(* IEC 61131-3 sources: plc-st-coding-agent/progress/f14_candidate/release/review/fixtures/agent_9772562, 4 files *)

(* ---- arm_one_step.st ---- *)
FUNCTION_BLOCK FB
VAR_INPUT
    ManualMode : BOOL;
    SingleStepMode : BOOL;
    SingleCycleMode : BOOL;
    ContinuousMode : BOOL;
    EmergencyStop : BOOL;
    Start : BOOL;
    DownButton : BOOL;
    UpButton : BOOL;
    LeftButton : BOOL;
    RightButton : BOOL;
    GripButton : BOOL;
    ReleaseButton : BOOL;
    DownLimitSwitch : BOOL;
    UpLimitSwitch : BOOL;
    LeftLimitSwitch : BOOL;
    RightLimitSwitch : BOOL;
    GripLimitSwitch : BOOL;
    ReleaseLimitSwitch : BOOL;
END_VAR
VAR_OUTPUT
    MoveDown : BOOL;
    MoveUp : BOOL;
    MoveLeft : BOOL;
    MoveRight : BOOL;
    ActivateGrip : BOOL;
    ActivateRelease : BOOL;
END_VAR
VAR
    step : INT := 1;
    busy : BOOL := FALSE;
    prevStart : BOOL := FALSE;
    prevManual : BOOL := FALSE;
    prevSingleStep : BOOL := FALSE;
    prevSingleCycle : BOOL := FALSE;
    prevContinuous : BOOL := FALSE;
    startRising : BOOL;
    autoSelected : BOOL;
    stepDone : BOOL;
END_VAR

(* 模式变化检测：任何模式输入改变时，停止当前动作并复位步骤 *)
IF (ManualMode <> prevManual) OR (SingleStepMode <> prevSingleStep) OR (SingleCycleMode <> prevSingleCycle) OR (ContinuousMode <> prevContinuous) THEN
    busy := FALSE;
    step := 1;
END_IF;
prevManual := ManualMode;
prevSingleStep := SingleStepMode;
prevSingleCycle := SingleCycleMode;
prevContinuous := ContinuousMode;

autoSelected := NOT ManualMode AND (SingleStepMode OR SingleCycleMode OR ContinuousMode);

startRising := Start AND NOT prevStart;
prevStart := Start;

IF autoSelected AND EmergencyStop THEN
    IF startRising THEN
        IF NOT busy THEN
            busy := TRUE;
        END_IF;
    END_IF;

    IF busy THEN
        stepDone := FALSE;
        CASE step OF
            1: stepDone := DownLimitSwitch;
            2: stepDone := GripLimitSwitch;
            3: stepDone := UpLimitSwitch;
            4: stepDone := RightLimitSwitch;
            5: stepDone := DownLimitSwitch;
            6: stepDone := ReleaseLimitSwitch;
            7: stepDone := UpLimitSwitch;
            8: stepDone := LeftLimitSwitch;
        END_CASE;

        IF stepDone THEN
            IF SingleStepMode THEN
                busy := FALSE;
                step := step MOD 8 + 1;
            ELSIF SingleCycleMode THEN
                IF step = 8 THEN
                    busy := FALSE;
                    step := 1;
                ELSE
                    step := step + 1;
                END_IF;
            ELSIF ContinuousMode THEN
                step := step MOD 8 + 1;
            END_IF;
        END_IF;
    END_IF;
END_IF;

IF EmergencyStop THEN
    IF ManualMode THEN
        MoveDown := DownButton AND NOT UpButton AND NOT DownLimitSwitch;
        MoveUp := UpButton AND NOT DownButton AND NOT UpLimitSwitch;
        MoveLeft := LeftButton AND NOT RightButton AND NOT LeftLimitSwitch;
        MoveRight := RightButton AND NOT LeftButton AND NOT RightLimitSwitch;
        ActivateGrip := GripButton AND NOT ReleaseButton AND NOT GripLimitSwitch;
        ActivateRelease := ReleaseButton AND NOT GripButton AND NOT ReleaseLimitSwitch;
    ELSIF autoSelected THEN
        IF busy THEN
            MoveDown := ((step = 1) OR (step = 5)) AND NOT DownLimitSwitch;
            MoveUp := ((step = 3) OR (step = 7)) AND NOT UpLimitSwitch;
            MoveLeft := (step = 8) AND NOT LeftLimitSwitch;
            MoveRight := (step = 4) AND NOT RightLimitSwitch;
            ActivateGrip := (step = 2) AND NOT GripLimitSwitch;
            ActivateRelease := (step = 6) AND NOT ReleaseLimitSwitch;
        ELSE
            MoveDown := FALSE;
            MoveUp := FALSE;
            MoveLeft := FALSE;
            MoveRight := FALSE;
            ActivateGrip := FALSE;
            ActivateRelease := FALSE;
        END_IF;
    ELSE
        MoveDown := FALSE;
        MoveUp := FALSE;
        MoveLeft := FALSE;
        MoveRight := FALSE;
        ActivateGrip := FALSE;
        ActivateRelease := FALSE;
    END_IF;
ELSE
    MoveDown := FALSE;
    MoveUp := FALSE;
    MoveLeft := FALSE;
    MoveRight := FALSE;
    ActivateGrip := FALSE;
    ActivateRelease := FALSE;
END_IF;

END_FUNCTION_BLOCK

(* ---- arm_restart.st ---- *)
FUNCTION_BLOCK FB
VAR_INPUT
    ManualMode : BOOL;
    SingleStepMode : BOOL;
    SingleCycleMode : BOOL;
    ContinuousMode : BOOL;
    EmergencyStop : BOOL;
    Start : BOOL;
    DownButton : BOOL;
    UpButton : BOOL;
    LeftButton : BOOL;
    RightButton : BOOL;
    GripButton : BOOL;
    ReleaseButton : BOOL;
    DownLimitSwitch : BOOL;
    UpLimitSwitch : BOOL;
    LeftLimitSwitch : BOOL;
    RightLimitSwitch : BOOL;
    GripLimitSwitch : BOOL;
    ReleaseLimitSwitch : BOOL;
END_VAR
VAR_OUTPUT
    MoveDown : BOOL;
    MoveUp : BOOL;
    MoveLeft : BOOL;
    MoveRight : BOOL;
    ActivateGrip : BOOL;
    ActivateRelease : BOOL;
END_VAR
VAR
    StartPrev : BOOL := FALSE;
    PrevManualMode : BOOL := FALSE;
    PrevSingleStepMode : BOOL := FALSE;
    PrevSingleCycleMode : BOOL := FALSE;
    PrevContinuousMode : BOOL := FALSE;
    ModeChanged : BOOL;
    StartPulse : BOOL;
    AutoStep : INT := 0;
END_VAR

MoveDown := FALSE;
MoveUp := FALSE;
MoveLeft := FALSE;
MoveRight := FALSE;
ActivateGrip := FALSE;
ActivateRelease := FALSE;

StartPulse := Start AND NOT StartPrev;
ModeChanged := (ManualMode <> PrevManualMode)
                OR (SingleStepMode <> PrevSingleStepMode)
                OR (SingleCycleMode <> PrevSingleCycleMode)
                OR (ContinuousMode <> PrevContinuousMode);

IF ModeChanged THEN
    AutoStep := 0;
END_IF;

IF EmergencyStop THEN
    IF ManualMode THEN
        MoveDown := DownButton AND NOT UpButton AND NOT DownLimitSwitch;
        MoveUp := UpButton AND NOT DownButton AND NOT UpLimitSwitch;
        MoveLeft := LeftButton AND NOT RightButton AND NOT LeftLimitSwitch;
        MoveRight := RightButton AND NOT LeftButton AND NOT RightLimitSwitch;
        ActivateGrip := GripButton AND NOT ReleaseButton AND NOT GripLimitSwitch;
        ActivateRelease := ReleaseButton AND NOT GripButton AND NOT ReleaseLimitSwitch;
    ELSIF SingleStepMode THEN
        IF AutoStep = 0 THEN
            IF StartPulse THEN
                AutoStep := 1;
            END_IF;
        END_IF;

        CASE AutoStep OF
            1:
                IF DownLimitSwitch THEN
                    AutoStep := 0;
                ELSE
                    MoveDown := TRUE;
                END_IF;
            2:
                IF GripLimitSwitch THEN
                    AutoStep := 0;
                ELSE
                    ActivateGrip := TRUE;
                END_IF;
            3:
                IF UpLimitSwitch THEN
                    AutoStep := 0;
                ELSE
                    MoveUp := TRUE;
                END_IF;
            4:
                IF RightLimitSwitch THEN
                    AutoStep := 0;
                ELSE
                    MoveRight := TRUE;
                END_IF;
            5:
                IF DownLimitSwitch THEN
                    AutoStep := 0;
                ELSE
                    MoveDown := TRUE;
                END_IF;
            6:
                IF ReleaseLimitSwitch THEN
                    AutoStep := 0;
                ELSE
                    ActivateRelease := TRUE;
                END_IF;
            7:
                IF UpLimitSwitch THEN
                    AutoStep := 0;
                ELSE
                    MoveUp := TRUE;
                END_IF;
            8:
                IF LeftLimitSwitch THEN
                    AutoStep := 0;
                ELSE
                    MoveLeft := TRUE;
                END_IF;
        END_CASE;
    ELSIF SingleCycleMode OR ContinuousMode THEN
        IF AutoStep = 0 THEN
            IF StartPulse THEN
                AutoStep := 1;
            END_IF;
        END_IF;

        IF AutoStep = 1 AND DownLimitSwitch THEN
            AutoStep := 2;
        END_IF;
        IF AutoStep = 2 AND GripLimitSwitch THEN
            AutoStep := 3;
        END_IF;
        IF AutoStep = 3 AND UpLimitSwitch THEN
            AutoStep := 4;
        END_IF;
        IF AutoStep = 4 AND RightLimitSwitch THEN
            AutoStep := 5;
        END_IF;
        IF AutoStep = 5 AND DownLimitSwitch THEN
            AutoStep := 6;
        END_IF;
        IF AutoStep = 6 AND ReleaseLimitSwitch THEN
            AutoStep := 7;
        END_IF;
        IF AutoStep = 7 AND UpLimitSwitch THEN
            AutoStep := 8;
        END_IF;
        IF AutoStep = 8 AND LeftLimitSwitch THEN
            IF ContinuousMode THEN
                AutoStep := 1;
            ELSE
                AutoStep := 0;
            END_IF;
        END_IF;

        CASE AutoStep OF
            1:
                IF NOT DownLimitSwitch THEN
                    MoveDown := TRUE;
                END_IF;
            2:
                IF NOT GripLimitSwitch THEN
                    ActivateGrip := TRUE;
                END_IF;
            3:
                IF NOT UpLimitSwitch THEN
                    MoveUp := TRUE;
                END_IF;
            4:
                IF NOT RightLimitSwitch THEN
                    MoveRight := TRUE;
                END_IF;
            5:
                IF NOT DownLimitSwitch THEN
                    MoveDown := TRUE;
                END_IF;
            6:
                IF NOT ReleaseLimitSwitch THEN
                    ActivateRelease := TRUE;
                END_IF;
            7:
                IF NOT UpLimitSwitch THEN
                    MoveUp := TRUE;
                END_IF;
            8:
                IF NOT LeftLimitSwitch THEN
                    MoveLeft := TRUE;
                END_IF;
        END_CASE;
    END_IF;
END_IF;

PrevManualMode := ManualMode;
PrevSingleStepMode := SingleStepMode;
PrevSingleCycleMode := SingleCycleMode;
PrevContinuousMode := ContinuousMode;
StartPrev := Start;
END_FUNCTION_BLOCK

(* ---- conveyor.st ---- *)
FUNCTION_BLOCK FB
VAR_INPUT
    processLength : USINT;
    sensor1 : BOOL;
    sensor2 : BOOL;
    sensor3 : BOOL;
    sensor4 : BOOL;
    sensor5 : BOOL;
    station1Start : BOOL;
    station2Complete : BOOL;
    station3Complete : BOOL;
    station4Complete : BOOL;
    processSequence : ARRAY[1..8] OF USINT;
END_VAR
VAR_OUTPUT
    conveyorLeft : BOOL;
    conveyorRight : BOOL;
END_VAR
VAR
    state : USINT := 0; (* 0=IDLE, 1=MOVING, 2=WAIT_PROCESS, 3=DONE *)
    currentStation : USINT := 1;
    seqIndex : USINT := 1;
    targetStation : USINT := 5;
    lastStation1Start : BOOL := FALSE;
    lastComplete2 : BOOL := FALSE;
    lastComplete3 : BOOL := FALSE;
    lastComplete4 : BOOL := FALSE;
END_VAR

(* 默认输出 *)
conveyorLeft := FALSE;
conveyorRight := FALSE;

(* 检查 processLength 有效性：若无效则强制停止并保持初始状态 *)
IF (processLength < 1) OR (processLength > 8) THEN
    state := 0;
    currentStation := 1;
    seqIndex := 1;
ELSE
    (* 状态机 *)
    IF (state = 0) OR (state = 3) THEN
        (* 启动检测：1# 传感器有料且启动按钮上升沿 *)
        IF (NOT lastStation1Start) AND station1Start AND sensor1 THEN
            seqIndex := 1;
            currentStation := 1;
            targetStation := processSequence[1];
            state := 1; (* MOVING *)
        END_IF
    ELSIF state = 1 THEN
        (* 移动中，检测目标传感器 *)
        IF (targetStation = 2) AND sensor2 THEN
            currentStation := 2;
            IF targetStation = 5 THEN
                state := 3; (* DONE *)
            ELSE
                state := 2; (* WAIT_PROCESS *)
            END_IF
        ELSIF (targetStation = 3) AND sensor3 THEN
            currentStation := 3;
            IF targetStation = 5 THEN
                state := 3;
            ELSE
                state := 2;
            END_IF
        ELSIF (targetStation = 4) AND sensor4 THEN
            currentStation := 4;
            IF targetStation = 5 THEN
                state := 3;
            ELSE
                state := 2;
            END_IF
        ELSIF (targetStation = 5) AND sensor5 THEN
            currentStation := 5;
            state := 3; (* DONE *)
        END_IF
    ELSIF state = 2 THEN
        (* 等待加工完成，检测对应完成信号上升沿 *)
        IF (currentStation = 2) AND (NOT lastComplete2) AND station2Complete THEN
            seqIndex := seqIndex + 1;
            IF seqIndex <= processLength THEN
                targetStation := processSequence[seqIndex];
                state := 1;
            ELSE
                state := 3;
            END_IF
        ELSIF (currentStation = 3) AND (NOT lastComplete3) AND station3Complete THEN
            seqIndex := seqIndex + 1;
            IF seqIndex <= processLength THEN
                targetStation := processSequence[seqIndex];
                state := 1;
            ELSE
                state := 3;
            END_IF
        ELSIF (currentStation = 4) AND (NOT lastComplete4) AND station4Complete THEN
            seqIndex := seqIndex + 1;
            IF seqIndex <= processLength THEN
                targetStation := processSequence[seqIndex];
                state := 1;
            ELSE
                state := 3;
            END_IF
        END_IF
    END_IF

    (* 设置输送方向输出 *)
    IF state = 1 THEN
        IF targetStation > currentStation THEN
            conveyorLeft := FALSE;
            conveyorRight := TRUE;
        ELSIF targetStation < currentStation THEN
            conveyorLeft := TRUE;
            conveyorRight := FALSE;
        ELSE
            conveyorLeft := FALSE;
            conveyorRight := FALSE;
        END_IF
    ELSE
        conveyorLeft := FALSE;
        conveyorRight := FALSE;
    END_IF
END_IF

(* 更新边沿历史 *)
lastStation1Start := station1Start;
lastComplete2 := station2Complete;
lastComplete3 := station3Complete;
lastComplete4 := station4Complete;

END_FUNCTION_BLOCK

(* ---- recipe.st ---- *)
TYPE ST_Recipe :
STRUCT
    recipeID : INT;
    ingredientType : INT;
    ingredientRatio : REAL;
    productionTemperature : REAL;
END_STRUCT
END_TYPE

FUNCTION_BLOCK FB
VAR_INPUT
    addRecipe : BOOL;
    deleteRecipe : BOOL;
    modifyRecipe : BOOL;
    queryRecipe : BOOL;
    recipeIn : ST_Recipe;
END_VAR
VAR_OUTPUT
    recipeAdded : BOOL;
    recipeDeleted : BOOL;
    recipeModified : BOOL;
    recipeQueryResult : ST_Recipe;
    error : BOOL;
    status : WORD;
END_VAR
VAR_IN_OUT
    recipe : ARRAY[1..10] OF ST_Recipe;
END_VAR
VAR
    prevAdd : BOOL := FALSE;
    prevDelete : BOOL := FALSE;
    prevModify : BOOL := FALSE;
    prevQuery : BOOL := FALSE;
    riseAdd : BOOL;
    riseDelete : BOOL;
    riseModify : BOOL;
    riseQuery : BOOL;
    i : INT;
    found : BOOL;
    emptyIndex : INT;
END_VAR

// 上升沿检测
riseAdd := addRecipe AND NOT prevAdd;
riseDelete := deleteRecipe AND NOT prevDelete;
riseModify := modifyRecipe AND NOT prevModify;
riseQuery := queryRecipe AND NOT prevQuery;

// 默认输出（无请求沿时保持）
recipeAdded := FALSE;
recipeDeleted := FALSE;
recipeModified := FALSE;
error := FALSE;
status := 0;

// 优先级：查询 > 添加 > 删除 > 修改
IF riseQuery THEN
    // 查询请求
    found := FALSE;
    FOR i := 1 TO 10 DO
        IF recipe[i].recipeID <> 0 AND recipe[i].recipeID = recipeIn.recipeID THEN
            recipeQueryResult := recipe[i];
            found := TRUE;
            EXIT;
        END_IF
    END_FOR
    IF NOT found THEN
        error := TRUE;
        status := 16#8001;
        // 清空查询结果
        recipeQueryResult.recipeID := 0;
        recipeQueryResult.ingredientType := 0;
        recipeQueryResult.ingredientRatio := 0.0;
        recipeQueryResult.productionTemperature := 0.0;
    END_IF
ELSIF riseAdd THEN
    // 添加请求
    found := FALSE;
    FOR i := 1 TO 10 DO
        IF recipe[i].recipeID <> 0 AND recipe[i].recipeID = recipeIn.recipeID THEN
            found := TRUE;
            EXIT;
        END_IF
    END_FOR
    IF found THEN
        error := TRUE;
        status := 16#8002;
    ELSE
        emptyIndex := 0;
        FOR i := 1 TO 10 DO
            IF recipe[i].recipeID = 0 THEN
                emptyIndex := i;
                EXIT;
            END_IF
        END_FOR
        IF emptyIndex = 0 THEN
            error := TRUE;
            status := 16#8003;
        ELSE
            recipe[emptyIndex] := recipeIn;
            recipeAdded := TRUE;
        END_IF
    END_IF
ELSIF riseDelete THEN
    // 删除请求
    found := FALSE;
    FOR i := 1 TO 10 DO
        IF recipe[i].recipeID <> 0 AND recipe[i].recipeID = recipeIn.recipeID THEN
            // 删除该槽，全部字段归零
            recipe[i].recipeID := 0;
            recipe[i].ingredientType := 0;
            recipe[i].ingredientRatio := 0.0;
            recipe[i].productionTemperature := 0.0;
            found := TRUE;
            EXIT;
        END_IF
    END_FOR
    IF found THEN
        recipeDeleted := TRUE;
    ELSE
        error := TRUE;
        status := 16#8004;
    END_IF
ELSIF riseModify THEN
    // 修改请求
    found := FALSE;
    FOR i := 1 TO 10 DO
        IF recipe[i].recipeID <> 0 AND recipe[i].recipeID = recipeIn.recipeID THEN
            recipe[i] := recipeIn;
            found := TRUE;
            EXIT;
        END_IF
    END_FOR
    IF found THEN
        recipeModified := TRUE;
    ELSE
        error := TRUE;
        status := 16#8005;
    END_IF
END_IF

// 更新上一周期信号
prevAdd := addRecipe;
prevDelete := deleteRecipe;
prevModify := modifyRecipe;
prevQuery := queryRecipe;

END_FUNCTION_BLOCK
